  # local inputrack = find_pattern_by_name("INPUT")
  # INSPECT_CONFIG_MAP.append(create_inspect_config(item_id=3, dx=inputrack.pattern_width[0]/(inputrack.pattern_size[0]-1), dy=inputrack.pattern_width[1]/(inputrack.pattern_size[1]-1), rack_size=inputrack.pattern_size , description="Input Capture"))
  # # Fills the Landmark List with Projectrelated Data
  # # create_landmark(lm_id=0, marker_id=-1, marker_size=0.1, marker_type="aruco_7x7", capture_pos=p[0,0,0,0,0,0], init_frame=p[0,0,0,0,0,0], search_offset=[0,0,0], actual_frame=p[0,0,0,0,0,0], description="")
  # LANDMARK_MAP.append(create_landmark(lm_id=1, marker_id=3, marker_size=0.1, marker_type="aruco_7x7", capture_pos = F10_Cap_CF, init_frame=p[-0.617789, -0.065471, 0.07918, 0.020983, -0.012695, 1.512066], search_offset=[0.15, 0.15, 0.1], actual_frame=p[-0.617789, -0.065471, 0.07918, 0.020983, -0.012695, 1.512066], description="LM CF Lid"))
  # LANDMARK_MAP.append(create_landmark(lm_id=2, marker_id=-1, marker_size=0.0085, marker_type="aruco_4x4", capture_pos = F8_Cap_Cobas_LM, init_frame=p[0,0,0,0,0,0], search_offset=[0.15, 0.15, 0.1], actual_frame=POS_Z, description="LM Cobas Rack Detection"))
  # LANDMARK_MAP.append(create_landmark(lm_id=3, marker_id=0, marker_size=0.1, marker_type="aruco_7x7", capture_pos = F17_Cobas_Cap, init_frame=p[-0.667,-0.194,0.100,0,0,0], search_offset=[0.15, 0.15, 0.1], actual_frame=POS_Z, description="LM Cobas Cap"))
  # LANDMARK_MAP.append(create_landmark(lm_id=4, marker_id=4, marker_size=0.1, marker_type="aruco_7x7", capture_pos = F19_XN550_Cap, init_frame=p[0.124,-0.976,0.355,-0.008,0.025,3.131], search_offset=[0.15, 0.15, 0.1], actual_frame=p[0,0,0,0,0,0], description="LM XN550 Cap"))
  # LANDMARK_MAP.append(create_landmark(lm_id=5, marker_id=0, marker_size=0.1, marker_type="aruco_7x7", capture_pos = TestLMCap, init_frame=p[-0.49,-0.144,0.092,0,-0.008,0.001], search_offset=[0.15, 0.15, 0.1], actual_frame=POS_Z, description="LM Test"))
  # # Configuration of all movement related parameters
  # # create_movement(id=0, hh_approach=POS_Z, h_approach=POS_Z, approach=POS_Z, h_target=POS_Z, target=POS_Z, retract=POS_Z, h_retract=POS_Z, hh_retract=POS_Z, h_frame=POS_Z, frame=POS_Z, speed=1, acceleration=1, description="default")
  # MOVEMENT_MAP.append(create_movement(description="TestLMCap", frame=TestLMCap, actionlist=[ActionManipulator.MOVE_TO]))
  # MOVEMENT_MAP.append(create_movement(description="TestLM", frame=TestLM, actionlist=[ActionManipulator.PICK,ActionManipulator.PLACE],
  #         approach=p[0,0,0.1,0,0,0],
  #         retract=p[0,0,0.1,0,0,0]))
  # MOVEMENT_MAP.append(create_movement(description="Home - MOVE_TO", frame=F1_uLM_Home, actionlist=[ActionManipulator.MOVE_TO]))
  # MOVEMENT_MAP.append(create_movement(description="Input - PICK&PLACE", frame=F2_uLM_Input, actionlist=[ActionManipulator.PICK,ActionManipulator.PLACE],
  #         approach=p[0,0,0.1,0,0,0],
  #         retract=p[0,0,0.1,0,0,0]))
  # MOVEMENT_MAP.append(create_movement(description="Capture Input - MOVE_TO", frame=F3_Cap_Input, actionlist=[ActionManipulator.MOVE_TO]))
  # MOVEMENT_MAP.append(create_movement(description="BIN - PLACE", frame=F4_uLM_Bin, actionlist=[ActionManipulator.PLACE],
  #         approach=p[0,0,0.1,0,0,0],
  #         retract=p[0,0,0.1,0,0,0]))
  # MOVEMENT_MAP.append(create_movement(description="Gripper - Move To", frame=F5_uLM_Gripper, actionlist=[ActionManipulator.MOVE_TO],
  #         approach=p[0,0,0.1,0,0,0]))
  # MOVEMENT_MAP.append(create_movement(description="Gripper - Pick", frame=F5_uLM_Gripper, actionlist=[ActionManipulator.PICK],
  #         retract=p[0,0,0.1,0,0,0]))
  # MOVEMENT_MAP.append(create_movement(description="Gripper - Place", frame=F5_uLM_Gripper, actionlist=[ActionManipulator.PLACE],
  #         approach=p[0,0,0.1,0,0,0]))
  # MOVEMENT_MAP.append(create_movement(description="CobasRack Pick & Place", frame=F6_uLM_Cobas_R, actionlist=[ActionManipulator.PICK,ActionManipulator.PLACE],
  #         approach=p[0,0,0.1,0,0,0],
  #         target=p[0,0,0,0,0,d2r(90)],
  #         retract=p[0,0,0.1,0,0,0]))
  # MOVEMENT_MAP.append(create_movement(description="CobasMagazine Pick & Place", frame=F7_uLM_Coba_Mag, actionlist=[ActionManipulator.PICK,ActionManipulator.PLACE],
  #         approach=p[0,0,0.1,0,0,0],
  #         target=p[0,0,0,0,0,-d2r(90)],
  #         retract=p[0,0,0.1,0,0,0]))
  # MOVEMENT_MAP.append(create_movement(description="Capture Position Cobas Landmarks", frame=F8_Cap_Cobas_LM, actionlist=[ActionManipulator.MOVE_TO]))
  # MOVEMENT_MAP.append(create_movement(description="TaraMagazine - PICK & PLACE", frame=F9_uLM_Tara, actionlist=[ActionManipulator.PICK,ActionManipulator.PLACE],
  #         approach=p[0,0,0.13,0,0,0],
  #         target=p[0,0,0,0,0,-d2r(90)],
  #         retract=p[0,0,0.13,0,0,0]))
  # MOVEMENT_MAP.append(create_movement(description="Capture Position - Centrifuge LM", frame=F10_Cap_CF,actionlist=[ActionManipulator.MOVE_TO]))
  # MOVEMENT_MAP.append(create_movement(description="Pick and Place Racks - Centrifuge Lid", frame=F11_CF_PiPl, actionlist=[ActionManipulator.PICK,ActionManipulator.PLACE],
  #         approach=p[0,0,0.3,0,0,0],
  #         retract=p[0,0,0.3,0,0,0]))
  # MOVEMENT_MAP.append(create_movement(description="Pick and Place Samples - Centrifuge on uLM", frame=F12_uLM_CF_Mag, actionlist=[ActionManipulator.PICK,ActionManipulator.PLACE],
  #         approach=p[0,0,0.13,0,0,0],
  #         retract=p[0,0,0.13,0,0,0]
  #         ))
  # MOVEMENT_MAP.append(create_movement(description="Pick and Place Racks - Centrifuge on uLM", frame=F13_uLM_CF_R, actionlist=[ActionManipulator.PICK,ActionManipulator.PLACE],
  #         approach=p[0,0,0.15,0,0,0],
  #         retract=p[0,0,0.15,0,0,0]
  #         ))

  # MOVEMENT_MAP.append(create_movement(description="Pick and Place Samples XN550 Racks in Device", frame=F18_XN550_Input, actionlist=[ActionManipulator.PICK,ActionManipulator.PLACE],
  #         approach=p[0,0,0.1,0,0,0],
  #         target = p[0,0,0,0,0,d2r(90)],
  #         retract=p[0,0,0.1,0,0,0]
  #         ))
  # MOVEMENT_MAP.append(create_movement(description="Capture LM XN550", frame=F19_XN550_Cap, actionlist=[ActionManipulator.MOVE_TO]))
  # MOVEMENT_MAP.append(create_movement(description="Open XN550 Drawer ", frame=F20_XN550_Draw, actionlist=[ActionManipulator.DRAWER_OPEN],
  #         h_approach=p[0.07,0,0.1,0,0,0],
  #         approach=p[0,0,0.1,0,0,0],
  #         target = p[0,0,0,0,0,d2r(90)],
  #         retract=p[0.07,0,0,0,0,0],
  #         h_retract=p[0.07,0,0.1,0,0,0]
  #         ))
  # MOVEMENT_MAP.append(create_movement(description="Close XN550 Drawer ", frame=F20_XN550_Draw, actionlist=[ActionManipulator.DRAWER_CLOSE],
  #         h_approach=p[0.07,0,0.1,0,0,0],
  #         approach=p[0.07,0,0,0,0,0],
  #         target = p[0,0,0,0,0,d2r(90)],
  #         retract=p[0,0,0.1,0,0,0],
  #         h_retract=p[0.07,0,0.1,0,0,0]
  #         ))
  # MOVEMENT_MAP.append(create_movement(description="Push XN550 Button ", frame=F21_XN550_Btn, actionlist=[ActionManipulator.PUSH],
  #         approach=p[0,0,0.15,0,0,0],
  #         retract=p[0,0,0.15,0,0,0]
  #         ))
  # MOVEMENT_MAP.append(create_movement(description="Capture Position 2 Input", frame=F_Cap_Input2,actionlist=[ActionManipulator.MOVE_TO]))



  $ 19 "Script: SCRIPT Objects V0.1.script"
  #*****************************************************
  # customer          :   INTERNAL
  # project name      :
  #****************************************************
  # controller        :   UR
  # software          :   5.17.3
  #****************************************************
  # author            :   P. Koehnke
  # Copyright (c)     :   United Robotics Group
  #                       An der Riede 2
  #                       28816 Stuhr
  #                       Germany
  #****************************************************
  # description       :   object database
  # version:      	:   0.1
  # created           :   09.10.2024
  # updated           :
  #****************************************************
  # modifications     :
  #
  # date              :
  # name              :
  # reason            :
  #****************************************************

  def create_object_2(id=0, name="", type=0, dimension=struct(length=0, width=0, height=0, diameter=0), gripper_offset=p[0,0,0,0,0,0]):
      return struct(id=id, name=name, type=type, dimension=dimension, gripper_offset=gripper_offset)
  end

  OBJ = create_object_2()
  OBJs = make_list(0, create_object_2(), 50)

  OBJs.append(create_object_2(id=1, name="rack centrifuge", type=1, dimension=struct(length=0, width=0, height=0.106, diameter=0.020), gripper_offset=p[0,0,0.095,0,0,2.356]))
  OBJs.append(create_object_2(id=2, name="sample tube 1", type=2, dimension=struct(length=0, width=0, height=0.106, diameter=0.015), gripper_offset=p[0,0,0,0,0,0]))
  OBJs.append(create_object_2(id=3, name="rack sarstedt", type=3, dimension=struct(length=0, width=0, height=0.100, diameter=0.020), gripper_offset=p[0,0,0,0,0,0]))
  OBJs.append(create_object_2(id=4, name="Lab bottle", type=4, dimension=struct(length=0, width=0, height=0.100, diameter=0.030), gripper_offset=p[0,0,0.2,0,0,0]))
  OBJs.append(create_object_2(id=5, name="Vial", type=5, dimension=struct(length=0, width=0, height=0.100, diameter=0.0275), gripper_offset=p[0,0,0,0,0,0]))
  OBJs.append(create_object_2(id=6, name="Container", type=6, dimension=struct(length=0.0, width=0.0, height=0, diameter=0.0), gripper_offset=p[0,0,0,0,0,0]))
  OBJs.append(create_object_2(id=7, name="Target_container", type=7, dimension=struct(length=0.06, width=0.06, height=0.134, diameter=0.05), gripper_offset=p[0,0,0,0,0,0]))
  OBJs.append(create_object_2(id=8, name="Spatula", type=8, dimension=struct(length=0.03, width=0.03, height=0.23, diameter=0.05), gripper_offset=p[0,0,0,0,0,0]))
  OBJs.append(create_object_2(id=9, name="rack pipet", type=9, dimension=struct(length=0.03, width=0.03, height=0.23, diameter=0.05), gripper_offset=p[0,0,0,0,0,0]))

  def create_jig_2(id=0, name="", type=0, capacity=0, jig_offset=p[0,0,0,0,0,0]):
      # iformation about used jigs
      return struct(id=id, name=name, type=type, capacity=capacity, jig_offset=jig_offset)
  end

  JIG2 = create_jig_2()
  JIGs = make_list(0, create_jig_2(), 20)

  JIGs.append(create_jig_2(id=1, name="3FG", type=1, capacity=1, jig_offset=p[0,0,0,0,0,0]))
  JIGs.append(create_jig_2(id=2, name="jig input", type=2, capacity=1, jig_offset=p[0,0,0,0,0,-3.927]))
  JIGs.append(create_jig_2(id=3, name="jig output", type=3, capacity=1, jig_offset=p[0,0,0,0,0,0.78]))
  JIGs.append(create_jig_2(id=6, name="jig bin", type=6, capacity=1, jig_offset=p[0,0,0,0,0,0]))
  JIGs.append(create_jig_2(id=7, name="jig sarstedt racks", type=7, capacity=1, jig_offset=p[0,0,-0.02,0,0,0]))
  JIGs.append(create_jig_2(id=8, name="NoK Bin", type=8, capacity=1, jig_offset=p[0,0,0,0,0,0]))
  JIGs.append(create_jig_2(id=9, name="Pick bott jig", type=9, capacity=1, jig_offset=p[0,0,0,0,0,0]))
  JIGs.append(create_jig_2(id=10, name="Place bott jig", type=10, capacity=1, jig_offset=p[0,0,0,0,0,0]))
  JIGs.append(create_jig_2(id=11, name="bottle shake jig", type=11, capacity=1, jig_offset=p[0,0,0,0,0,0]))
  JIGs.append(create_jig_2(id=12, name="Pick Vial jig", type=12, capacity=1, jig_offset=p[0,0,0,0,0,0]))
  JIGs.append(create_jig_2(id=13, name="Place Vial jig", type=13, capacity=1, jig_offset=p[0,0,0,0,0,0]))
  JIGs.append(create_jig_2(id=14, name="Liquid transfer jig", type=14, capacity=1, jig_offset=p[0,0,0,0,0,0]))
  JIGs.append(create_jig_2(id=15, name="Pick station jig", type=15, capacity=1, jig_offset=p[0,0,0,0,0,0]))
  JIGs.append(create_jig_2(id=16, name="Place station jig", type=16, capacity=1, jig_offset=p[0,0,0,0,0,0]))
  JIGs.append(create_jig_2(id=17, name="Weigh station jig", type=17, capacity=1, jig_offset=p[0,0,0,0,0,0]))
  JIGs.append(create_jig_2(id=18, name="Pick station 1", type=18, capacity=1, jig_offset=p[0,0,0,0,0,0]))
  JIGs.append(create_jig_2(id=19, name="Pick station 2", type=19, capacity=1, jig_offset=p[0,0,0,0,0,0]))
  JIGs.append(create_jig_2(id=20, name="Pick station 3", type=20, capacity=1, jig_offset=p[0,0,0,0,0,0]))
  JIGs.append(create_jig_2(id=21, name="Tilt station jig", type=21, capacity=1, jig_offset=p[0,0,0,0,0,0]))
  $ 26 "Script: Powder_all.script"
  global SERVER_IP   = "192.168.12.139"
  global SERVER_PORT = 3002

  global container_id = 0
  global powder_id  = 0
  global bulk_density = 0
  global H          = 0
  global H_c          = 0
  global mouth_d     = 0
  global mouth_sh    = 0
  global length_c     = 0
  global diameter   = 0
  global empty_weight_g  = 0
  global volume_ml    = 0
  global shape_code   = 0
  global flow_code   = 0
  global shape = ""
  global Flowability = ""
  global full_weight_g = 0
  global cent_edge = 0
  global pick_2_base = 0.2 # distance from tcp to base of picking table
  global wall_thickness = 0.001

  def read_db_data():

    socket_open(SERVER_IP, SERVER_PORT)
    sleep(0.5)
    socket_send_string("GET_DATACODE_FLOATS")
    sleep(5)

    local fl = socket_read_ascii_float(14)
    socket_close()

    global container_id = fl[1]
    global powder_id = fl[2]
    global bulk_density = fl[3]
    global H          = fl[4]/1000
    global H_c          = fl[5]/1000
    global mouth_d     = fl[6]/1000
    global mouth_sh    = fl[7]/1000
    global length_c     = fl[8]/1000
    global diameter   = fl[9]/1000
    global empty_weight_g = fl[10]
    global volume_ml    = fl[11]
    global full_weight_g = fl[12]
    global flow_code   = fl[13]
    global shape_code   = fl[14]

  	if (flow_code == 1.0):
  	  global Flowability = "MEDIUM"
  	elif (flow_code == 2.0):
  	  global Flowability = "LOW"
  	else:
  	  global Flowability = "HIGH"
  	end

    if ( shape_code == 1.0):
  	shape = "cylindrical"
  	cent_edge =  diameter
    else:
  	shape = "cubical"
  	cent_edge =  length_c
    end

  end


  def send_picking_info(Pow_name, target_weight):
    socket_open(SERVER_IP, SERVER_PORT)
    cmd = "PICK:"+Pow_name+";"+to_str(target_weight)
    socket_send_string(cmd)
    sleep(0.1)
    socket_close()
  end

  #### POTS ####
  def tilt_send(angle):
  	socket_open("192.168.12.101", 80)
  	angle = 90.0 - angle
  	socket_send_string("Tilt,"+to_str(angle)+",0")
  	sync()
  	sleep(0.5)
  	socket_close()
  end

  def Motors_off():
  	socket_open("192.168.12.101", 80)
  	socket_send_string("Off,0,0")
  	sync()
  	sleep(0.5)
  	socket_close()
  end

  def Rotate():
  	socket_open("192.168.12.101", 80)
  	socket_send_string("FullRotation, 1, 2000")
  	sync()
  	sleep(0.5)
  	socket_close()
  end

  def CCW_Rotate():
  	socket_open("192.168.12.101", 80)
  	socket_send_string("FullRotation, -1, 2000")
  	sync()
  	sleep(0.5)
  	socket_close()
  end

  def tilt_to_home():
  	socket_open("192.168.12.101", 80)
  	socket_send_string("Home,0,0")
  	sync()
  	sleep(0.5)
  	socket_close()
  end
  #######
  def vibration_1():
  	set_analog_out(0,0.4)
  	sleep(1)
  	set_analog_out(0,0.0)
  	sleep(0)
  end

  def vibration_2():
  	set_analog_out(0,0.4)
  	sleep(0.8)
  	set_analog_out(0,0.0)
  	sleep(0.2)
  end

  def vibration_3():
  	set_analog_out(0,0.4)
  	sleep(0.5)
  	set_analog_out(0,0.0)
  	sleep(0.3)
  end

  def vibration_4():
  	set_analog_out(0,0.8)
  	sleep(0.6)
  	set_analog_out(0, 0.0)
  	sleep(0.5)
  end

  ##################

  global gear_2_holder = 0.018
  global gain_per_percent = 0.5
  global w_dosed_total = 0.0
  global last_scale = 0.0
  global tilt_angle_sent = 0.0
  global level = 0.0
  global target_g = 0.0
  global angle_max = 60
  global angle_min = 10
  global hinge_2_base = 0.0421
  global TCP_2_tip_x = 0.0047
  global spatula_len = 0.182
  global spatula_offset = p[TCP_2_tip_x,0,spatula_len,0,0,0]
  global SPATULA_L_VOL_ML = 5.0        # 1 teaspoon = 5 mL
  global SPATULA_M_VOL_ML = 1.25       # 1/4 teaspoon = 1.25 mL
  global SPATULA_S_VOL_ML = 0.15625    # 1/32 teaspoon = 0.15625 mL
  global SPATULA_FLAT_M_VOL_ML  = 2.2
  global SPATULA_FLAT_S_VOL_ML  = 1.2   #based on caluclations using rho = m/V
  global ry_deg_safe = 0
  global ry_deg = 0



  def clamp(x, lo, hi):
  	if(x<lo):
  		return lo
  	elif (x>hi):
  		return hi
  	else:
  		return x
  	end
  end

  def compute_level_percent(W_now, weight_value):   # W_now = container+powder, weight_value = live scale reading
      local delta = weight_value - last_scale

      if (delta < 0.0):
          delta = 0.0
      end

      global w_dosed_total = w_dosed_total + delta
      global last_scale = weight_value     # update the last scale reading

      local W_eff = W_now - w_dosed_total
      if (W_eff <  empty_weight_g):
          W_eff =  empty_weight_g
      end

      # Compute powder level %
      level = 100.0 * (W_eff -  empty_weight_g) / (full_weight_g -  empty_weight_g)

      # Clamp to 0–100
      level = clamp(level, 0, 100)
    textmsg("deb 1 = ", level)
      return level
  end

  def deg2rad(d):
  	return d*3.141592/180
  end

  def my_abs(val):
  	if (val<0):
  		return -val
  	else:
  		return val
  	end
  end

  def compute_tilt_deg(level_percent):
  	angle = angle_min + gain_per_percent*(100.0-level_percent)

    	textmsg("deb 2 = ", angle)
  	return clamp(angle, angle_min, angle_max)
  end

  def tilt(level_percentage):
  	new_angle = compute_tilt_deg(level_percentage)
  	global angle_rel = new_angle - tilt_angle_sent

  	if my_abs(angle_rel)>2.0:
  		tilt_send(new_angle)
  		global angle_deg = new_angle
  		global tilt_angle_sent = new_angle
  		global p_center_vertical = center_pose()
  		global p_center = updated_center_pose(p_center_vertical, angle_deg)
  	end

  	if (level_percentage<85.0):
  		tilt_send(angle_deg)
  	end
  end

  def compute_scoop_depth(level):
    return ((100.0-level)/100.0)*(H -mouth_sh )
  end

  def map_tilt_to_ry_deg(container_deg, level):

  	if (Flowability == "HIGH" or Flowability == "MEDIUM"):
  		global scoop_depth = compute_scoop_depth(level)
  		safe_scoop_pivot = (mouth_d  - spatula_depth)/(scoop_depth+mouth_sh )
  		global ry_deg_safe = asin(safe_scoop_pivot)
  		global ry_deg = 90-container_deg
  	else:
  		global scoop_depth = compute_scoop_depth(level)
  		safe_scoop_pivot = (mouth_d  - spatula_depth)/(scoop_depth+mouth_sh )
  		global ry_deg_safe = asin(safe_scoop_pivot)
  		global ry_deg = 90-container_deg
  	end
  	return [ry_deg_safe,ry_deg]
  end

  def get_scoop_weight(spatula, bulk_density):

  	local vol = 0

  	if (spatula == "spatula_L"):
  		vol = SPATULA_L_VOL_ML
  		global spatula_depth = 0.015
  		global spatula_mid   = 0.016
  		global spatula_ry    = 0.0

  	elif (spatula == "spatula_M"):
  		vol = SPATULA_M_VOL_ML
  		global spatula_depth = 0.010
  		global spatula_mid   = 0.0105
  		global spatula_ry    = 0.0

  	elif (spatula == "spatula_S"):
  		vol = SPATULA_S_VOL_ML
  		global spatula_depth = 0.008
  		global spatula_mid   = 0.0063
  		global spatula_ry    = 0.0

  	elif (spatula == "spatula_flat_M"):
  		vol = SPATULA_FLAT_M_VOL_ML
  		global spatula_depth = 0.001
  		global spatula_mid   = 0.002
  		global spatula_ry    = 10.0

  	elif (spatula == "spatula_flat_S"):
  		vol = SPATULA_FLAT_S_VOL_ML
  		global spatula_depth = 0.005
  		global spatula_mid   = 0.016
  		global spatula_ry    = 2.0

  	else:
  		textmsg("Unknown spatula type")
  		return 0.0
  	end
  	global target_g = vol * bulk_density
  	return target_g

  end

  def select_spatula(Flowability, level, diff, bulk_density, mouth_d ):

      local k = 1.1

      global powder_height = (H  - mouth_sh ) * level/100

      # =====================================================
      # LOW FLOWABILITY
      # =====================================================
      if (Flowability == "LOW"):

          local gFM = get_scoop_weight("spatula_flat_M", bulk_density)

          local level_ok_FM = (spatula_mid * 2 < powder_height)
          local diff_ok_FM  = (diff > k * gFM)

          local flatM_ok = level_ok_FM and diff_ok_FM

          if (flatM_ok):
              return "spatula_flat_M"
          else:
              return "spatula_flat_S"
          end

      end


      # =====================================================
      # LARGE
      # =====================================================
      local gL = get_scoop_weight("spatula_L", bulk_density)

      local mouth_ok_L = (mouth_d  >= 0.05)
      local level_ok_L = (spatula_mid * 2 < powder_height)
      local diff_ok_L  = (diff > k * gL)

      local large_ok = mouth_ok_L and level_ok_L and diff_ok_L


      # =====================================================
      # MEDIUM
      # =====================================================
      local gM = get_scoop_weight("spatula_M", bulk_density)

      local level_ok_M = (spatula_mid * 2 < powder_height)
      local diff_ok_M  = (diff > k * gM)

      local medium_ok = level_ok_M and diff_ok_M


      # =====================================================
      # FINAL SELECTION
      # =====================================================
      if (large_ok):
          return "spatula_L"

      elif (medium_ok):
          return "spatula_M"

      else:
          return "spatula_S"
      end

  end

  def after_scoop():
  	tilt_send(angle_deg)
  	sleep(0.5)
  	movel(lifted_pose, a=0.05, v=0.2)
  	movel(tilted_pose_in_base2, a=0.05, v=0.2)
  	set_analog_out(0,0.4)
  	movel(pose_trans(tilted_pose_in_base2, p[0,0,0,0,0,2.0]), a=0.05, v=0.2)
  	set_analog_out(0,0.0)
  	movel(lifted_pose, a=0.05, v=0.2)
  	tilt_to_home()
  end

  def center_pose():
  	global p_translated = container_place
  	#global p_translated = pots_axis_temp

  	#cx = p_translated[0]
  	#cy = p_translated[1]
  	#cz = p_translated[2]

  	global p_center_vertical_temp = pose_trans(p_translated, p[0,0,0, deg2rad(90), 0, 0])
  	cx = p_center_vertical_temp[0]
  	cy = p_center_vertical_temp[1]
  	cz = p_center_vertical_temp[2]
  	#rx = p_center_vertical_temp[3]
  	#ry = p_center_vertical_temp[4]
  	rz = p_center_vertical_temp[5]

  	global p_center_vertical_temp = p[cx,cy,cz, 0, 0, rz]
  	trans_rel = p[0,0,-pick_2_base+H,0,0,0]
  	global p_center_vertical =  pose_trans(p_center_vertical_temp, trans_rel)
  	return p_center_vertical
  end

  def updated_center_pose(p_center_vertical, angle_deg):
  	hinge_pose = pose_trans(p_center_vertical, p[0,0,-hinge_2_base-gear_2_holder-H ,0,0,0])
  	local_rel = pose_trans(pose_inv(hinge_pose), p_center_vertical)

  	rot_tilt = p[0,0,0, -deg2rad(angle_deg),0,0]
  	local_rel_tilted = pose_trans(rot_tilt, local_rel)

  	global p_center = pose_trans(hinge_pose, local_rel_tilted)
  	return p_center
  end

  def scoop_powder(p_center):
  	vibration_voltage = 0.4
  	vibration_time = 3.0
  	global scoop_radius_default = 0.0


  	scoop_radius_default = mouth_d /2 - spatula_depth
  	scoop_safe_entry_pose = pose_trans(p_center, p[-TCP_2_tip_x,0,spatula_len+0.05,0,0,0])
  	scoop_entry_pose = pose_trans(p_center, p[-TCP_2_tip_x,0,spatula_len,0,0,0])

  	movel(scoop_safe_entry_pose, a=0.1, v=0.25)
  	movel(scoop_entry_pose, a=0.1, v=0.25)

  	scoop_start_rel_int = p[0, 0, -mouth_sh , 0, 0, 0]
  	scoop_start_pose_int = pose_trans(scoop_entry_pose, scoop_start_rel_int)

  	movel(scoop_start_pose_int, a=0.1, v=0.25)

  	if (spatula_mid * 2 < powder_height and spatula == "spatula_M" or spatula == "spatula_L"):

  		global total_depth = mouth_sh + scoop_depth + spatula_mid
  		global total_depth = clamp(total_depth, 0, H - spatula_mid)
  		scoop_start_rel = p[scoop_radius_default, 0, -total_depth, 0, 0, 0]

  		rot_mid = p[0, 0, 0, 0, 0, 0.785]
  		rot_end = p[0, 0, 0, 0, 0, 1.5708]

  		scoop_via_rel = pose_trans(rot_mid, scoop_start_rel)
  		scoop_end_rel = pose_trans(rot_end, scoop_start_rel)

  		scoop_start_pose = pose_trans(scoop_entry_pose, scoop_start_rel)
  		scoop_via_pose = pose_trans(scoop_entry_pose, scoop_via_rel)
  		scoop_end_pose = pose_trans(scoop_entry_pose, scoop_end_rel)

  		movel(scoop_start_pose, a=0.5, v=0.3)

  		if (level<90.0):
  			Rotate()
  		end

  		movec(scoop_via_pose, scoop_end_pose, a=0.03, v=0.02)
  		sleep(1.0)
  		#local ry_deg = map_tilt_to_ry_deg(angle_deg,level)
  		local ry_result = map_tilt_to_ry_deg(angle_deg,level)
  		global ry_safe = ry_result[0]
  		global ry = deg2rad(ry_result[1])

  		# safe_retention
  		local pivot_pose = pose_trans(scoop_end_pose, p[0,0,total_depth-spatula_len,0,0,0])
  		local end_rel = pose_trans(pose_inv(pivot_pose), scoop_end_pose)
  		local end_rel_tilted = pose_trans(end_rel, p[0, 0, 0, 0, ry_safe, 0])
  		global tilted_pose_in_base = pose_trans(pivot_pose, p[0,0,0,end_rel_tilted[3],end_rel_tilted[4], end_rel_tilted[5]])
  		global tilted_pose_in_base = pose_trans(tilted_pose_in_base, p[0, 0, spatula_len-total_depth, 0, 0, 0])
  		# sptula pivoted around the container rim of the mouth at ry_safe
  		movel(tilted_pose_in_base, a=0.03, v=0.1)

  		#popup("is the spatula crashing at front? ", blocking = True)
  		# safe_retention_above
  		# calculate x , z movements

  		global safe_x = sin(ry_safe)*(scoop_depth - (mouth_d -spatula_depth)/tan(90-ry_safe/2))
  		global safe_z = cos(ry_safe)*(scoop_depth - (mouth_d -spatula_depth)/tan(90-ry_safe/2))

  		local safe_up = pose_trans(tilted_pose_in_base, p[-safe_x,0,safe_z,0,0,0])
  		movel(safe_up, a=0.03, v=0.1)

  		#popup("is the spatula crashing at neck? ", blocking = True)

  		# full exit step by step
  		#local alpha = atan(2*mouth_sh /mouth_d )

  		#global cent_pose_cont_x = sin(ry_safe)*(scoop_depth - (mouth_d -spatula_depth)/tan(90-ry_safe/2))
  		#global cent_pose_cont_z = cos(ry_safe)*(scoop_depth+mouth_sh  - (mouth_d -spatula_depth)/tan(90-ry_safe/2))
  		#local cent_pose_cont = pose_trans(safe_up, p[])

  		# full exit
  		local pivot_pose2 = pose_trans(tilted_pose_in_base, p[0,0,total_depth-spatula_len,0,0,0])
  		local end_rel2 = pose_trans(pose_inv(pivot_pose2), tilted_pose_in_base)
  		#popup("is the spatula crashing front? ", blocking = True)
  		local end_rel_tilted2 = pose_trans(end_rel2, p[0, 0, 0, 0, ry-ry_safe, 0])
  		global tilted_pose_in_base2 = pose_trans(pivot_pose2, p[0,0,0,end_rel_tilted2[3],end_rel_tilted2[4], end_rel_tilted2[5]])
  		global tilted_pose_in_base2 = pose_trans(tilted_pose_in_base2, p[-TCP_2_tip_x, 0, spatula_len-scoop_radius_default-spatula_mid, 0, 0, 0])
  		# spaula exited at center of the mouth at ry
  		movel(tilted_pose_in_base2, a=0.03, v=0.1)
  		#popup("is the spatula crashing at mouth? ", blocking = True)

  	else : # emptying logic
  		spatula_base = pose_trans(scoop_entry_pose, p[0, 0, -H, 0, 0, 0])
  		local pivot_pose = pose_trans(scoop_entry_pose, p[0,0,-spatula_len,0,0,0])
  		# tilt inwards
  		global in_angle = atan((cent_edge-spatula_depth)/(2*H))
  		spatula_tilt_rel = pose_trans(pose_inv(pivot_pose), spatula_base)

  		spatula_tilt = pose_trans(spatula_tilt_rel, p[0, 0, 0, in_angle, 0, 0])
  		global tilted_pose = pose_trans(pivot_pose, p[0,0,0,spatula_tilt[3],spatula_tilt[4], spatula_tilt[5]])

  		global tilted_pose = pose_trans(tilted_pose, p[0,0,spatula_len-H,0,0,0])

  		movel(tilted_pose,a=0.1, v=0.25)
  		Rotate()

  		rot_mid = p[0, 0, 0, 0, 0, 0.785]
  		rot_end = p[0, 0, 0, 0, 0, 1.5708]

  		scoop_via_rel = pose_trans(tilted_pose, rot_mid)
  		scoop_end_rel = pose_trans(tilted_pose, rot_end)

  		movec(scoop_via_rel, scoop_end_rel, a=0.03, v=0.02)
  		popup("is the spatula crashing front? ", blocking = True)

  		scoop_via_pose = pose_trans(pivot_pose, scoop_via_rel)
  		scoop_end_pose = pose_trans(pivot_pose, scoop_end_rel)

  		#movec(scoop_via_pose, scoop_end_pose, a=0.03, v=0.02)
  		popup("is the spatula crashing front? ", blocking = True)
  		local ry_result = map_tilt_to_ry_deg(angle_deg,level)
  		global ry_safe = ry_result[0]
  		global ry = deg2rad(ry_result[1])

  		# full exit
  		#local pivot_pose2 = pose_trans(scoop_entry_pose, p[0,0,-spatula_len,0,0,0])
  		local end_rel2 = pose_trans(pose_inv(pivot_pose), scoop_end_pose)
  		popup("is the spatula crashing front? ", blocking = True)
  		local end_rel_tilted2 = pose_trans(end_rel2, p[0, 0, 0, 0, ry, 0])
  		global tilted_pose_in_base2 = pose_trans(pivot_pose, p[0,0,0,end_rel_tilted2[3],end_rel_tilted2[4], end_rel_tilted2[5]])
  		global tilted_pose_in_base2 = pose_trans(tilted_pose_in_base2, p[0, 0, spatula_len, 0, 0, 0])
  		# sptula exited at center of the mouth at ry
  		movel(tilted_pose_in_base2, a=0.03, v=0.1)
  		popup("is the spatula crashing at mouth? ", blocking = True)
  	end

  	if (spatula=="spatula_flat_S" or spatula=="spatula_S"):
  		vibration_3()
  	elif (spatula == "spatula_M"):
  		vibration_4()
  	else:
  		set_analog_out(0, vibration_voltage)
  	end

  	# remove excess
  	local pivot_pose_level = pose_trans(tilted_pose_in_base2, p[0,0,-spatula_len,0,0,0])
  	local end_rel_level = pose_trans(pose_inv(pivot_pose_level), tilted_pose_in_base2)
  	#local ry_level = ry/1.5
  	local ry_level = deg2rad(15)
  	local end_rel_tilted_level = pose_trans(end_rel_level, p[0, 0, 0, 0, -ry_level, 0])
  	local end_rel_tilted_level2 = pose_trans(pivot_pose_level, p[0, 0, 0,end_rel_tilted_level[3],end_rel_tilted_level[4], end_rel_tilted_level[5]])
  	local end_rel_tilted_level2 = pose_trans(end_rel_tilted_level2, p[0,0,spatula_len,0,0,0])
  	movel(end_rel_tilted_level2, a=0.03, v=0.1)

  	movel(tilted_pose_in_base2, a=0.03, v=0.1)
  	set_analog_out(0, 0.0)
  	#popup("safe out + moving towards beaker", title = "Pause", blocking = True)
  	global lifted_pose = pose_trans(tilted_pose_in_base2, p[-0.04,0,0.04,0,0,0]) # safety distance away from the container

  	movel(lifted_pose, a=0.03, v=0.1)
  	CCW_Rotate()
  end

  def auto_tilt_and_scoop(W_now, target_weight, weight_value):
  	global level = compute_level_percent(W_now, weight_value)

  	global spatula = select_spatula(Flowability, level, diff, bulk_density, mouth_d )
  	textmsg("deb 4 8 = ", spatula)
  	#global target_g = get_scoop_weight(spatula, bulk_density)

    	#textmsg("deb 4 = ", target_g)
  	#send_scoop_target_info()

  	global scoop_depth = compute_scoop_depth(level)

    	textmsg("deb 5 = ", scoop_depth)
  	tilt_to_home()
  	sleep(0.5)
  	tilt(level)
  	sleep(1.5)
    	#popup("is the pots tilted? ", blocking = True)
    	#textmsg("deb 6 = ", p_center)
  	scoop_powder(p_center)

    	textmsg("deb 7 - sucess")
  end
  $ 27 "Script: Weight_scale_socket_s.script"
  global s_depth = 0
  global s_length =0
  global s_volume = 0
  global ry_theta  = 0

  def get_weight():
  	socket_open(SERVER_IP,SERVER_PORT)
  	sleep(0.2)
  	textmsg("socket opened successfully!")
  	socket_send_string("GET_WEIGHT")
  	sleep(0.2)
  	sync()
  	sleep(0.2)
  	receiveFromServ = socket_read_ascii_float(6)
  	sleep(1)
  	#while (receiveFromServ[0] <1):
  		#receiveFromServ = socket_read_ascii_float(1)
  		#sleep(1)
  		#textmsg("retrying read:", receiveFromServ)
  	#end
  	textmsg("Received weight:", receiveFromServ[1])
  	sleep(0.2)
  	socket_close()
  	sleep(0.2)
  	return receiveFromServ[1]
  end

  def tare_scale():
  	socket_open(SERVER_IP,SERVER_PORT)
  	socket_send_string("TARE")
  	sleep(2)
  	socket_close()
  end

  def zero_scale():
  	socket_open(SERVER_IP,SERVER_PORT)
  	socket_send_string("ZERO")
  	sleep(0.5)
  	socket_close()
  end

  def log_weight():
  	socket_open(SERVER_IP,SERVER_PORT)
  	socket_send_string("LOG_WEIGHT")
  	sleep(0.5)
  	socket_close()
  end

  def send_target_info():
  	socket_open(SERVER_IP,SERVER_PORT)
  	socket_send_string("SET_TARGET:" + to_str(target_weight))
  	sleep(0.2)
  	socket_close()
  end
  def send_powder_info():
  	socket_open(SERVER_IP,SERVER_PORT)
  	socket_send_string("SET_POWDER:" + Pow_name)
  	sleep(0.2)
  	socket_close()
  end
  def send_spatula_info():
  	socket_open(SERVER_IP,SERVER_PORT)
  	socket_send_string("SET_SPATULA:" + spatula)
  	#sleep(1)

  	#local fl = socket_read_ascii_float(4)
    	#socket_close()

    	#global s_depth = fl[1]
    	#global s_length = fl[2]
   	#global s_volume = fl[3]
   	#global ry_theta  = fl[4]
  	sleep(0.2)

  end

  def send_level_info():
  	socket_open(SERVER_IP,SERVER_PORT)
  	socket_send_string("SET_LEVEL:" + to_str(level))
  	sleep(0.2)
  	socket_close()
  end
  def send_weight_info():
    socket_open(SERVER_IP, SERVER_PORT)
    #rq_open_and_wait()
    cmd = "GET_CONT_WEIGHT"
    socket_send_string(cmd)
    sync()
    sleep(0.5)
    receiveFromSer = socket_read_ascii_float(1)
    socket_close()
    return receiveFromSer[1]
  end

  $ 28 "BeforeStarts"
  $ 29 "uLM"
  $ 30 "CMD_Stop≔ False "
  global CMD_Stop=  False
  $ 31 "CMD_Abort≔ False "
  global CMD_Abort=  False
  $ 32 "CMD_Clear≔ False "
  global CMD_Clear=  False
  $ 33 "STATE≔1"
  global STATE=1
  $ 34 "STATE_Info≔''"
  global STATE_Info=""
  $ 35 "ARM_Referenced≔ False "
  global ARM_Referenced=  False
  $ 36 "zero_ftsensor()"
  zero_ftsensor()
  $ 37 "poses init"
  $ 38 "PSE_A≔p[0,0,0,0,0,0]"
  global PSE_A=p[0,0,0,0,0,0]
  $ 39 "PSE_A_H≔p[0,0,0,0,0,0]"
  global PSE_A_H=p[0,0,0,0,0,0]
  $ 40 "PSE_R≔p[0,0,0,0,0,0]"
  global PSE_R=p[0,0,0,0,0,0]
  $ 41 "PSE_R_H≔p[0,0,0,0,0,0]"
  global PSE_R_H=p[0,0,0,0,0,0]
  $ 42 "PSE_T≔p[0,0,0,0,0,0]"
  global PSE_T=p[0,0,0,0,0,0]
  $ 43 "PSE_T_H≔p[0,0,0,0,0,0]"
  global PSE_T_H=p[0,0,0,0,0,0]
  $ 44 "PSE_C_E≔p[0,0,0,0,0,0]"
  global PSE_C_E=p[0,0,0,0,0,0]
  $ 45 "PSE_C_H≔p[0,0,0,0,0,0]"
  global PSE_C_H=p[0,0,0,0,0,0]
  $ 46 "PSE_C_S≔p[0,0,0,0,0,0]"
  global PSE_C_S=p[0,0,0,0,0,0]
  $ 47 "init_home_by_cartesian_pose(p[0,-0.400,0.300,0,0,0])"
  init_home_by_cartesian_pose(p[0,-0.400,0.300,0,0,0])
  $ 48 "Clearing"
  $ 49 "reset_error()"
  reset_error()
  $ 50 "reset_warning()"
  reset_warning()
  $ 51 "uGo"
  $ 53 "ugo_init( True ,'http://192.168.12.120:10001')"
  ugo_init(  True  ,"http://192.168.12.120:10001")
  $ 54 "ugo_update_outputs()"
  ugo_update_outputs()
  $ 55 "App"
  $ 56 "'ADD APPLICATION SPECIFIC COMMANDS'"
  # 'ADD APPLICATION SPECIFIC COMMANDS'
  $ 57 "Tools"
  $ 58 "OBJ_Picked≔gripper_has_object()"
  global OBJ_Picked=gripper_has_object()
  $ 59 "If OBJ_Picked"
  if (OBJ_Picked):
    # begin: URCap Program Node
    #   Source: Robotiq_Grippers, 3.17.0.105337, Robotiq Inc.
    #   Type: Gripper Activate
    $ 60 "Gripper Activate"

    kill rq_gripper_communication_thread
    rq_gripper_communication_thread_started = False
    rq_close_gripper_socket("1")
    rq_close_gripper_socket("2")
    rq_close_gripper_socket("3")
    rq_close_gripper_socket("4")

    rq_init_comm_if_connected(9, "1")
    rq_init_comm_if_connected(2, "2")
    rq_init_comm_if_connected(3, "3")
    rq_init_comm_if_connected(4, "4")
    rq_print_connected_grippers()
    rq_gripper_communication_thread = run rq_gripper_communication()

    while(not rq_gripper_communication_thread_started):
        sleep(0.008)
    end

    rq_set_max_current_for_all_grippers()

    reset_and_activate = False

    rq_activate_all_grippers(False)
    # end: URCap Program Node
  else:
    $ 61 "Else" "noBreak"
    # begin: URCap Program Node
    #   Source: Robotiq_Grippers, 3.17.0.105337, Robotiq Inc.
    #   Type: Gripper Activate
    $ 62 "Gripper Reset and Activate"

    kill rq_gripper_communication_thread
    rq_gripper_communication_thread_started = False
    rq_close_gripper_socket("1")
    rq_close_gripper_socket("2")
    rq_close_gripper_socket("3")
    rq_close_gripper_socket("4")

    rq_init_comm_if_connected(9, "1")
    rq_init_comm_if_connected(2, "2")
    rq_init_comm_if_connected(3, "3")
    rq_init_comm_if_connected(4, "4")
    rq_print_connected_grippers()
    rq_gripper_communication_thread = run rq_gripper_communication()

    while(not rq_gripper_communication_thread_started):
        sleep(0.008)
    end

    rq_set_max_current_for_all_grippers()

    reset_and_activate = True

    rq_activate_all_grippers(True)
    # end: URCap Program Node
  end
  $ 63 "zero_ftsensor()"
  zero_ftsensor()
  $ 64 "EXTT"
  $ 65 "Set GRP_3F_Enable=Off"
  set_standard_digital_out(4, False)
  $ 66 "Set BarcodeTrigger=Off"
  set_standard_digital_out(6, False)
  $ 67 "Set GRP_3F_Decap=Off"
  set_standard_digital_out(3, False)
  $ 68 "Set GRP_3F_Cap=Off"
  set_standard_digital_out(2, False)
  $ 69 "Set GRP_3F_Open=Off"
  set_standard_digital_out(5, False)
  $ 70 "PSE_T≔get_tool_free_pose(dir=[0,0,0.150], move_in_base_frame=True)"
  global PSE_T=get_tool_free_pose(dir=[0,0,0.150], move_in_base_frame=True)
  $ 71 "If is_reachable(Base_const, [PSE_T])"
  if (is_reachable(p[0.0,0.0,0.0,0.0,0.0,0.0], [PSE_T])):
    $ 72 "MoveL"
    $ 73 "PSE_T" "breakAfter"
    movel(PSE_T, a=1.2, v=0.15)
  end
  $ 75 "powder dispensing variable init"
  $ 76 "Start_thread≔ False "
  global Start_thread=  False
  $ 77 "vib_thread≔ False "
  global vib_thread=  False
  $ 78 "QR assignment init"
  $ 79 "d_cc≔0.06"
  global d_cc=0.06
  $ 81 "kp≔0.0015"
  global kp=0.0015
  $ 82 "ki≔0.0001"
  global ki=0.0001
  $ 83 "kd≔0.01"
  global kd=0.01
  $ 84 "dt≔0.03"
  global dt=0.03
  $ 85 "Integral_error≔0"
  global Integral_error=0
  $ 86 "current_error≔0"
  global current_error=0
  $ 87 "previous_error≔0"
  global previous_error=0
  $ 88 "tilt_increment≔0"
  global tilt_increment=0
  $ 89 "tilt_angle≔0"
  global tilt_angle=0
  $ 90 "diff≔0"
  global diff=0
  $ 91 "current_pose≔get_actual_tcp_pose()"
  global current_pose= get_actual_tcp_pose ()
  $ 92 "Relative_trans≔p[0, 0, -0.035, 0, 0, 0]"
  global Relative_trans=p[0, 0, -0.035, 0, 0, 0]
  $ 96 "tilt_to_home()"
  tilt_to_home()
  $ 97 "switch_spat_M≔ True "
  global switch_spat_M=  True
  $ 98 "switch_spat_S≔ True "
  global switch_spat_S=  True
  $ 99 "switch_spat_F_M≔ True "
  global switch_spat_F_M=  True
  $ 100 "switch_spat_F_S≔ True "
  global switch_spat_F_S=  True
  $ 101 "last_scale≔0"
  global last_scale=0
  $ 793 "Thread_1"
  thread Thread_1():
    while (True):
      $ 794 "If Start_thread≟ True "
      if (Start_thread ==   True  ):
        $ 795 "weight_value≔get_weight()"
        global weight_value=get_weight()
        $ 796 "Wait: 0.2"
        sleep(0.2)
        $ 797 "sync()"
        sync()
      end
      $ 798 "sync()"
      sync()
    end
  end
  threadId_Thread_1 = run Thread_1()
  $ 799 "Thread_2"
  thread Thread_2():
    while (True):
      $ 800 "Loop vib_thread≟ True "
      thread Thread_while_800():
        while (True):
          $ 801 "diff≔target_weight-weight_value"
          global diff=target_weight-weight_value
          $ 802 "If diff>0.02 and spatula≠'spatula_flat_S'"
          global thread_flag_802=0
          thread Thread_if_802():
            $ 804 "Set AO[0]=4.0"
            set_standard_analog_out(0, 0.4)
            thread_flag_802 = 1
          end
          if (diff>0.02  and  spatula != "spatula_flat_S"):
            global thread_handler_802=run Thread_if_802()
            while (thread_flag_802 == 0):
              if not(diff>0.02  and  spatula != "spatula_flat_S"):
                kill thread_handler_802
                thread_flag_802 = 2
              else:
                sync()
              end
            end
          else:
            thread_flag_802 = 2
          end
          if (thread_flag_802 == 2):
            $ 805 "ElseIf diff>0.02 and spatula≟'spatula_flat_S'"
            if (diff>0.02 and spatula == "spatula_flat_S"):
              $ 806 "vibration_3()"
              vibration_3()
            else:
              $ 807 "ElseIf diff≤0.03"
              global thread_flag_807=0
              thread Thread_if_807():
                $ 808 "vibration_2()"
                vibration_2()
                thread_flag_807 = 1
              end
              if (diff <= 0.03):
                global thread_handler_807=run Thread_if_807()
                while (thread_flag_807 == 0):
                  if not(diff <= 0.03):
                    kill thread_handler_807
                    thread_flag_807 = 2
                  else:
                    sync()
                  end
                end
              else:
                thread_flag_807 = 2
              end
              if (thread_flag_807 == 2):
                $ 813 "Else" "noBreak"
                $ 814 "Set AO[0]=0.0"
                set_standard_analog_out(0, 0.0)
              end
            end
          end
        end
      end
      if (vib_thread ==   True  ):
        global thread_handler_800=run Thread_while_800()
        while (vib_thread ==   True  ):
          sync()
        end
        kill thread_handler_800
      end
      $ 815 "sync()"
      sync()
    end
  end
  threadId_Thread_2 = run Thread_2()
  while (True):
    $ 102 "Robot Program"
    $ 103 "MAIN"
    $ 104 "command_manager(external_control='uGO', cond_suspend=(ITM_Manipulated and AMR_AtTarget and AMR_Charging and AMR_Battery<40), cond_unsuspend=(AMR_Battery≟60))"
    command_manager(external_control="uGO", cond_suspend=(ITM_Manipulated  and  AMR_AtTarget  and  AMR_Charging  and  AMR_Battery<40), cond_unsuspend=(AMR_Battery == 60))
    $ 105 "log_state(STATE_Info)"
    log_state(STATE_Info)
    $ 106 "Switch STATE"
    switch_1 = STATE
    $ 107 "Case 1"
    if (1 == switch_1):
      $ 108 "Stopping"
      $ 109 "STATE_Info≔'Stopping'"
      global STATE_Info="Stopping"
      $ 110 "end_freedrive_mode()"
      end_freedrive_mode()
      $ 111 "Set"
      set_tcp(p[0.0,0.0,0.161,3.1415,0.0,0.0])
      $ 112 "PSE_T≔get_tool_free_pose(dir=[0,0,0.150], move_in_base_frame=True)"
      global PSE_T=get_tool_free_pose(dir=[0,0,0.150], move_in_base_frame=True)
      $ 113 "If is_reachable(Base_const, [PSE_T])"
      if (is_reachable(p[0.0,0.0,0.0,0.0,0.0,0.0], [PSE_T])):
        $ 114 "MoveL"
        $ 115 "PSE_T" "breakAfter"
        movel(PSE_T, a=1.2, v=0.15)
      end
      $ 116 "do_transition(keep_rxry=OBJ_Picked, r=0)"
      do_transition(keep_rxry=OBJ_Picked, r=0)
      $ 125 "Call Sub_AMR_MiR_V3"
      Sub_AMR_MiR_V3()
      $ 126 "If stopping() and AMR_Done"
      if (stopping()  and  AMR_Done):
        $ 127 "STATE≔2"
        global STATE=2
        $ 128 "ugo_update_outputs()"
        ugo_update_outputs()
      end
    elif (2 == switch_1):
      $ 129 "Case 2"
      $ 130 "Stopped"
      $ 131 "STATE_Info≔'Stopped'"
      global STATE_Info="Stopped"
      $ 132 "Call Sub_AMR_MiR_V3"
      Sub_AMR_MiR_V3()
      $ 133 "If CMD_Reset  or PB_Start"
      if (CMD_Reset   or  get_standard_digital_in(0)):
        $ 134 "STATE≔3"
        global STATE=3
        $ 135 "ugo_update_outputs()"
        ugo_update_outputs()
      end
    elif (3 == switch_1):
      $ 136 "Case 3"
      $ 137 " Resetting"
      $ 138 "STATE_Info≔'Resetting'"
      global STATE_Info="Resetting"
      $ 139 "uML"
      $ 140 "reset_error()"
      reset_error()
      $ 141 "reset_warning()"
      reset_warning()
      $ 142 "PROCESS_Step≔0"
      global PROCESS_Step=0
      $ 143 "PROCESS_Info≔''"
      global PROCESS_Info=""
      $ 144 "ARM_Referenced≔ False "
      global ARM_Referenced=  False
      $ 145 "WRK_Done≔ False "
      global WRK_Done=  False
      $ 146 "ITM_Prepared≔ False "
      global ITM_Prepared=  False
      $ 147 "ITM_Manipulated≔ False "
      global ITM_Manipulated=  False
      $ 148 "STP≔0"
      global STP=0
      $ 149 "Action≔0"
      global Action=0
      $ 150 "Action_Info≔''"
      global Action_Info=""
      $ 151 "ITM_ID≔0"
      global ITM_ID=0
      $ 152 "JIG≔0"
      global JIG=0
      $ 153 "JIG_Slot≔0"
      global JIG_Slot=0
      $ 154 "Task_info≔''"
      global Task_info=""
      $ 155 "Set"
      set_tcp(p[0.0,0.0,0.161,3.1415,0.0,0.0])
      $ 156 "App"
      $ 157 "'ADD APPLICATION SPECIFIC COMMANDS'"
      # 'ADD APPLICATION SPECIFIC COMMANDS'
      $ 158 "OBJ_Type≔0"
      global OBJ_Type=0
      $ 159 "OBJ_Nbr≔0"
      global OBJ_Nbr=0
      $ 160 "If CNT_Rack_Output≥50"
      if (CNT_Rack_Output >= 50):
        $ 161 "CNT_Rack_Output≔0"
        global CNT_Rack_Output=0
      end
      $ 162 "TASK≔struct(ID=0, NAVI=struct(target=0, footprint=0, protectiveOff=0, dock=0), WORK=struct(ITM_ID_Src=0, JIG_ID_Src=0, OBJ_Nbr_Src=0, ACT_Src=0, ITM_ID_Tgt=0, JIG_ID_Tgt=0, OBJ_Nbr_Tgt=0, ACT_Tgt=0, OBJ_Type=0))"
      global TASK=struct(ID=0, NAVI=struct(target=0, footprint=0, protectiveOff=0, dock=0), WORK=struct(ITM_ID_Src=0, JIG_ID_Src=0, OBJ_Nbr_Src=0, ACT_Src=0, ITM_ID_Tgt=0, JIG_ID_Tgt=0, OBJ_Nbr_Tgt=0, ACT_Tgt=0, OBJ_Type=0))
      $ 163 "Call Sub_AMR_MiR_V3"
      Sub_AMR_MiR_V3()
      $ 164 "If resetting() and AMR_Done"
      if (resetting()  and  AMR_Done):
        $ 165 "STATE≔4"
        global STATE=4
        $ 166 "ugo_update_outputs()"
        ugo_update_outputs()
      end
    elif (4 == switch_1):
      $ 167 "Case 4"
      $ 168 "Idle"
      $ 169 "STATE_Info≔'Idle'"
      global STATE_Info="Idle"
      $ 170 "If CMD_Start"
      if (CMD_Start):
        $ 171 "STATE≔5"
        global STATE=5
        $ 172 "ugo_update_outputs()"
        ugo_update_outputs()
      end
    elif (5 == switch_1):
      $ 173 "Case 5"
      $ 174 "Starting"
      $ 175 "STATE_Info≔'Starting'"
      global STATE_Info="Starting"
      $ 176 "'ADD COMMANDS WHAT TO START WITH'"
      # 'ADD COMMANDS WHAT TO START WITH'
      $ 177 "Call Sub_AMR_MiR_V3"
      Sub_AMR_MiR_V3()
      $ 178 "get ugo data"
      $ 179 "Assign Tasks"
      $ 180 "TASK.ID = ugo_get_task()"
      TASK.ID = ugo_get_task()
      $ 181 "If TASK.ID≟1"
      if (TASK.ID == 1):
        $ 182 "Task_info≔'Charge'"
        global Task_info="Charge"
        $ 183 "Parameters"
        $ 184 "AMR_PosTarget≔1"
        global AMR_PosTarget=1
      else:
        $ 185 "ElseIf TASK.ID≟9"
        if (TASK.ID == 9):
          $ 186 "'Pick Sarstedt Rack from Variable source'"
          # 'Pick Sarstedt Rack from Variable source'
          $ 187 "Task_info≔'Navigate to Target'"
          global Task_info="Navigate to Target"
          $ 188 "Parameters"
          $ 189 "AMR_PosTarget≔UGO.read_input('00','ITM_ID')"
          global AMR_PosTarget=UGO.read_input("00","ITM_ID")
        else:
          $ 190 "ElseIf TASK.ID≟13"
          if (TASK.ID == 13):
            $ 191 "Task_info≔'Dose Powder'"
            global Task_info="Dose Powder"
            $ 192 "Parameters"
            $ 193 "ITM_ID≔1"
            global ITM_ID=1
            $ 194 "W_now≔(UGO.read_input('00','Container_weight'))/1000"
            global W_now=(UGO.read_input("00","Container_weight"))/1000
            $ 195 "Pow_name≔(UGO.read_input('00','Powder_name'))"
            global Pow_name=(UGO.read_input("00","Powder_name"))
            $ 196 "target_weight≔(UGO.read_input('00','Target_weight'))/1000"
            global target_weight=(UGO.read_input("00","Target_weight"))/1000
            $ 197 "send_picking_info(Pow_name,target_weight)"
            send_picking_info(Pow_name,target_weight)
            $ 198 "OBJ_Type≔6"
            global OBJ_Type=6
            $ 199 "JIG≔17"
            global JIG=17
            $ 200 "AMR_PosTarget≔5"
            global AMR_PosTarget=5
          else:
            $ 201 "ElseIf TASK.ID≟49"
            if (TASK.ID == 49):
              $ 202 "Task_info≔'Pick Containers'"
              global Task_info="Pick Containers"
              $ 203 "Parameters"
              $ 204 "ITM_ID≔1"
              global ITM_ID=1
              $ 205 "OBJ_Type≔6"
              global OBJ_Type=6
              $ 206 "JIG≔15"
              global JIG=15
              $ 207 "AMR_PosTarget≔3"
              global AMR_PosTarget=3
            else:
              $ 208 "ElseIf TASK.ID≟50"
              if (TASK.ID == 50):
                $ 209 "Task_info≔'Decap Containers'"
                global Task_info="Decap Containers"
                $ 210 "Parameters"
                $ 211 "ITM_ID≔1"
                global ITM_ID=1
                $ 212 "OBJ_Type≔6"
                global OBJ_Type=6
                $ 213 "JIG≔16"
                global JIG=16
                $ 214 "AMR_PosTarget≔5"
                global AMR_PosTarget=5
              else:
                $ 215 "ElseIf TASK.ID≟51"
                if (TASK.ID == 51):
                  $ 216 "Task_info≔'Detect Spatula and transfer powder'"
                  global Task_info="Detect Spatula and transfer powder"
                  $ 217 "Parameters"
                  $ 218 "ITM_ID≔1"
                  global ITM_ID=1
                  $ 219 "target_weight≔(UGO.read_input('00','Target_weight'))/1000"
                  global target_weight=(UGO.read_input("00","Target_weight"))/1000
                  $ 220 "OBJ_Type≔8"
                  global OBJ_Type=8
                  $ 221 "JIG≔16"
                  global JIG=16
                  $ 222 "AMR_PosTarget≔5"
                  global AMR_PosTarget=5
                else:
                  $ 223 "ElseIf TASK.ID≟52"
                  if (TASK.ID == 52):
                    $ 224 "Task_info≔'Pick Powder'"
                    global Task_info="Pick Powder"
                    $ 225 "Parameters"
                    $ 226 "ITM_ID≔1"
                    global ITM_ID=1
                    $ 228 "OBJ_Type≔6"
                    global OBJ_Type=6
                    $ 229 "JIG≔15"
                    global JIG=15
                    $ 230 "AMR_PosTarget≔3"
                    global AMR_PosTarget=3
                  else:
                    $ 231 "ElseIf TASK.ID≟53"
                    if (TASK.ID == 53):
                      $ 232 "Task_info≔'Decap Powder'"
                      global Task_info="Decap Powder"
                      $ 233 "Parameters"
                      $ 234 "ITM_ID≔1"
                      global ITM_ID=1
                      $ 235 "OBJ_Type≔6"
                      global OBJ_Type=6
                      $ 236 "JIG≔1"
                      global JIG=1
                      $ 237 "AMR_PosTarget≔5"
                      global AMR_PosTarget=5
                    else:
                      $ 238 "ElseIf TASK.ID≟54"
                      if (TASK.ID == 54):
                        $ 239 "Task_info≔'Empty and swap Powder container'"
                        global Task_info="Empty and swap Powder container"
                        $ 248 "Parameters"
                        $ 249 "ITM_ID≔1"
                        global ITM_ID=1
                        $ 251 "W_now≔(UGO.read_input('00','Container_weight'))/1000"
                        global W_now=(UGO.read_input("00","Container_weight"))/1000
                        $ 252 "Pow_name≔(UGO.read_input('00','Powder_name'))"
                        global Pow_name=(UGO.read_input("00","Powder_name"))
                        $ 255 "OBJ_Type≔6"
                        global OBJ_Type=6
                        $ 256 "JIG≔17"
                        global JIG=17
                        $ 257 "AMR_PosTarget≔5"
                        global AMR_PosTarget=5
                      else:
                        $ 258 "ElseIf TASK.ID≟55"
                        if (TASK.ID == 55):
                          $ 259 "Task_info≔'Place Powder'"
                          global Task_info="Place Powder"
                          $ 260 "Parameters"
                          $ 261 "ITM_ID≔1"
                          global ITM_ID=1
                          $ 262 "OBJ_Type≔6"
                          global OBJ_Type=6
                          $ 263 "JIG≔21"
                          global JIG=21
                          $ 264 "AMR_PosTarget≔5"
                          global AMR_PosTarget=5
                        else:
                          $ 265 "ElseIf TASK.ID≟56"
                          if (TASK.ID == 56):
                            $ 266 "Task_info≔'Dose Powder'"
                            global Task_info="Dose Powder"
                            $ 267 "Parameters"
                            $ 268 "ITM_ID≔1"
                            global ITM_ID=1
                            $ 269 "target_weight≔(UGO.read_input('00','Target_weight'))/1000"
                            global target_weight=(UGO.read_input("00","Target_weight"))/1000
                            $ 270 "W_now≔(UGO.read_input('00','Container_weight'))/1000"
                            global W_now=(UGO.read_input("00","Container_weight"))/1000
                            $ 271 "Pow_name≔(UGO.read_input('00','Powder_name'))"
                            global Pow_name=(UGO.read_input("00","Powder_name"))
                            $ 272 "OBJ_Type≔6"
                            global OBJ_Type=6
                            $ 273 "JIG≔17"
                            global JIG=17
                            $ 274 "AMR_PosTarget≔5"
                            global AMR_PosTarget=5
                          else:
                            $ 275 "ElseIf TASK.ID≟57"
                            if (TASK.ID == 57):
                              $ 276 "Task_info≔'Recipe Powder dosing'"
                              global Task_info="Recipe Powder dosing"
                              $ 277 "Parameters"
                              $ 278 "ITM_ID≔1"
                              global ITM_ID=1
                              $ 279 "Pow_A≔(UGO.read_input('00','PowderA'))"
                              global Pow_A=(UGO.read_input("00","PowderA"))
                              $ 280 "Pow_B≔(UGO.read_input('00','PowderB'))"
                              global Pow_B=(UGO.read_input("00","PowderB"))
                              $ 281 "Pow_C≔(UGO.read_input('00','PowderC'))"
                              global Pow_C=(UGO.read_input("00","PowderC"))
                              $ 282 "Total_weight≔(UGO.read_input('00','Total_weight'))/1000"
                              global Total_weight=(UGO.read_input("00","Total_weight"))/1000
                              $ 283 "Pow_A_percent≔(UGO.read_input('00','PowderA_percentage'))/100"
                              global Pow_A_percent=(UGO.read_input("00","PowderA_percentage"))/100
                              $ 284 "Pow_B_percent≔(UGO.read_input('00','PowderB_percentage'))/100"
                              global Pow_B_percent=(UGO.read_input("00","PowderB_percentage"))/100
                              $ 285 "Pow_C_percent≔(UGO.read_input('00','PowderC_percentage'))/100"
                              global Pow_C_percent=(UGO.read_input("00","PowderC_percentage"))/100
                              $ 286 "OBJ_Type≔6"
                              global OBJ_Type=6
                              $ 287 "JIG≔17"
                              global JIG=17
                              $ 288 "AMR_PosTarget≔5"
                              global AMR_PosTarget=5
                            else:
                              $ 289 "ElseIf TASK.ID≟58"
                              if (TASK.ID == 58):
                                $ 290 "Task_info≔'Pick Powder containers'"
                                global Task_info="Pick Powder containers"
                                $ 291 "Parameters"
                                $ 292 "ITM_ID≔1"
                                global ITM_ID=1
                                $ 293 "OBJ_Type≔6"
                                global OBJ_Type=6
                                $ 294 "JIG≔15"
                                global JIG=15
                                $ 295 "AMR_PosTarget≔3"
                                global AMR_PosTarget=3
                              else:
                                $ 296 "Else" "noBreak"
                                $ 297 "set_error(ERROR_WRONG_ORDER)"
                                set_error(ERROR_WRONG_ORDER)
                              end
                            end
                          end
                        end
                      end
                    end
                  end
                end
              end
            end
          end
        end
      end
      $ 298 "test ugo"
      $ 299 "Wait: 0.2"
      sleep(0.2)
      $ 300 "ugo_update_outputs()"
      ugo_update_outputs()
      $ 301 "If starting() and AMR_Done"
      if (starting()  and  AMR_Done):
        $ 302 "log_message(Task_info, 'New Task: ')"
        log_message(Task_info, "New Task: ")
        $ 303 "log_message(to_str(TASK.ID), 'Task_ID: ')"
        log_message(to_str(TASK.ID), "Task_ID: ")
        $ 304 "do_transition(keep_rxry=OBJ_Picked)"
        do_transition(keep_rxry=OBJ_Picked)
        $ 305 "STATE≔6"
        global STATE=6
        $ 306 "ugo_update_outputs()"
        ugo_update_outputs()
      end
    elif (6 == switch_1):
      $ 307 "Case 6"
      $ 308 "Execute"
      $ 309 "STATE_Info≔'Execute'"
      global STATE_Info="Execute"
      $ 310 "If  not CMD_Hold and not CMD_Suspend"
      global thread_flag_310=0
      thread Thread_if_310():
        $ 311 "Switch PROCESS_Step"
        switch_2 = PROCESS_Step
        $ 312 "Case 0"
        if (0 == switch_2):
          $ 313 "PROCESS_Info≔'process control'"
          global PROCESS_Info="process control"
          $ 314 "log_process(PROCESS_Info)"
          log_process(PROCESS_Info)
          $ 315 "process control"
          $ 316 "If  not AMR_AtTarget"
          if (  not  AMR_AtTarget):
            $ 317 "PROCESS_Step≔1"
            global PROCESS_Step=1
          else:
            $ 318 "ElseIf (( not ITM_Prepared and  not WRK_Done) or (ITM_Prepared and WRK_Done))"
            if (((  not  ITM_Prepared  and    not  WRK_Done)  or  (ITM_Prepared  and  WRK_Done))):
              $ 319 "PROCESS_Step≔2"
              global PROCESS_Step=2
            else:
              $ 320 "ElseIf  not WRK_Done"
              if (  not  WRK_Done):
                $ 321 "PROCESS_Step≔3"
                global PROCESS_Step=3
              else:
                $ 322 "Else" "noBreak"
                $ 323 "task finished"
                $ 324 "PROCESS_Info≔''"
                global PROCESS_Info=""
                $ 325 "STATE≔7"
                global STATE=7
                $ 326 "ugo_update_outputs()"
                ugo_update_outputs()
              end
            end
          end
        elif (1 == switch_2):
          $ 327 "Case 1"
          $ 328 "navigate"
          $ 329 "'MOVING THE uML'"
          # 'MOVING THE uML'
          $ 330 "PROCESS_Info≔'move to target'"
          global PROCESS_Info="move to target"
          $ 331 "log_process(PROCESS_Info)"
          log_process(PROCESS_Info)
          $ 332 "If TASK.ID≟1"
          if (TASK.ID == 1):
            $ 333 "Action≔51"
            global Action=51
          else:
            $ 334 "Else" "noBreak"
            $ 335 "Action≔52"
            global Action=52
          end
          $ 336 "Call Sub_AMR_MiR_V3"
          Sub_AMR_MiR_V3()
          $ 337 "If AMR_Done"
          if (AMR_Done):
            $ 338 "PROCESS_Step≔0"
            global PROCESS_Step=0
          end
        elif (2 == switch_2):
          $ 339 "Case 2"
          $ 340 "prepare"
          $ 341 "'THINGS THAT HAVE TO BE DONE ONCE IN A SEQUENCE,WORKFLOW'"
          # 'THINGS THAT HAVE TO BE DONE ONCE IN A SEQUENCE,WORKFLOW'
          $ 342 "PROCESS_Info≔'prepare for work'"
          global PROCESS_Info="prepare for work"
          $ 343 "log_process(PROCESS_Info)"
          log_process(PROCESS_Info)
          $ 344 "If TASK.WORK.ITM_ID_Src>1"
          if (TASK.WORK.ITM_ID_Src>1):
            $ 345 "ITM_ID≔TASK.WORK.ITM_ID_Src"
            global ITM_ID=TASK.WORK.ITM_ID_Src
          else:
            $ 346 "ElseIf TASK.WORK.ITM_ID_Tgt>1"
            if (TASK.WORK.ITM_ID_Tgt>1):
              $ 347 "ITM_ID≔TASK.WORK.ITM_ID_Tgt"
              global ITM_ID=TASK.WORK.ITM_ID_Tgt
            end
          end
          $ 348 "If  not ARM_Referenced and (ITM_ID≠0)"
          if (  not  ARM_Referenced  and  (ITM_ID != 0)):
            $ 349 "STP≔1"
            global STP=1
          else:
            $ 350 "ElseIf ARM_Referenced or (ITM_ID≟0)"
            if (ARM_Referenced  or  (ITM_ID == 0)):
              $ 351 "STP≔2"
              global STP=2
            end
          end
          $ 352 "Switch STP"
          switch_3 = STP
          $ 353 "Case 1"
          if (1 == switch_3):
            $ 354 "reference"
            $ 355 "STP_Info≔'reference at target position'"
            global STP_Info="reference at target position"
            $ 356 "log_step(STP_Info)"
            log_step(STP_Info)
            $ 357 "If ITM_ID≟1"
            if (ITM_ID == 1):
              $ 358 "CAM_Done≔ True "
              global CAM_Done=  True
            else:
              $ 359 "Else" "noBreak"
              $ 360 "Action≔131"
              global Action=131
              $ 361 "Call Sub_Vision_V18"
              Sub_Vision_V18()
            end
            $ 363 "If CAM_Done and  not ERROR.FLAG"
            if (CAM_Done  and    not  ERROR.FLAG):
              $ 364 "log_step('ARM referenced')"
              log_step("ARM referenced")
              $ 365 "ARM_Referenced≔ True "
              global ARM_Referenced=  True
            end
          elif (2 == switch_3):
            $ 366 "Case 2"
            $ 367 "manipulate"
            $ 368 "STP_Info≔'manipulate item'"
            global STP_Info="manipulate item"
            $ 369 "log_step(STP_Info)"
            log_step(STP_Info)
            $ 370 "'In case pressing button is needed'"
            # 'In case pressing button is needed'
            $ 371 "If found_in_list(ITM_ID, ITM_ID_List)"
            if (found_in_list(ITM_ID, ITM_ID_List)):
              $ 372 "Switch ITM_ID"
              switch_4 = ITM_ID
              $ 373 "Case 0"
              if (0 == switch_4):
                $ 374 "ITM_Manipulated≔ not ITM_Manipulated"
                global ITM_Manipulated=  not  ITM_Manipulated
              elif (1 == switch_4):
                $ 375 "Case 1"
                $ 376 "ITM_Manipulated≔ not ITM_Manipulated"
                global ITM_Manipulated=  not  ITM_Manipulated
              elif (2 == switch_4):
                $ 377 "Case 2"
              else:
                $ 387 "Default Case"
                $ 388 "ITM_Manipulated≔ not ITM_Manipulated"
                global ITM_Manipulated=  not  ITM_Manipulated
              end
            end
          end
          $ 389 "ITM_Prepared≔(ITM_Manipulated or  not found_in_list(ITM_ID, ITM_ID_List)) and (ARM_Referenced or ITM_ID≟0) and  not WRK_Done"
          global ITM_Prepared=(ITM_Manipulated  or    not  found_in_list(ITM_ID, ITM_ID_List))  and  (ARM_Referenced  or  ITM_ID == 0)  and    not  WRK_Done
          $ 390 "STP≔0"
          global STP=0
          $ 391 "STP_Info≔''"
          global STP_Info=""
          $ 392 "PROCESS_Step≔0"
          global PROCESS_Step=0
        elif (3 == switch_2):
          $ 393 "Case 3"
          $ 394 "work"
          $ 395 "'ADD EVERY MACHINE, OBJECT, STATION TO WORK ON'"
          # 'ADD EVERY MACHINE, OBJECT, STATION TO WORK ON'
          $ 396 "Switch ITM_ID"
          switch_3 = ITM_ID
          $ 397 "Case 1"
          if (1 == switch_3):
            $ 398 "uLM"
            $ 399 "If TASK.ID≟12"
            if (TASK.ID == 12):
              $ 400 "fill racks"
              $ 401 "Action≔151"
              global Action=151
              $ 402 "Call Sub_Vision_V18"
              Sub_Vision_V18()
              $ 403 "If  not ERROR.FLAG"
              if (  not  ERROR.FLAG):
                $ 404 "Actions for the task"
                $ 405 "Action≔1"
                global Action=1
                $ 406 "JIG≔2"
                global JIG=2
                $ 407 "JIG_Slot≔CAM_Result[0]"
                global JIG_Slot=CAM_Result[0]
                $ 408 "OBJ_Nbr≔CAM_Result[0]"
                global OBJ_Nbr=CAM_Result[0]
                $ 409 "OBJ_Type≔2"
                global OBJ_Type=2
                $ 410 "Call Sub_Action_V4"
                Sub_Action_V4()
                $ 411 "If OBJ_Picked"
                if (OBJ_Picked):
                  $ 412 "CAM_Result.remove(0)"
                  CAM_Result.remove(0)
                  $ 413 "PRC_TubCounter≔PRC_TubCounter+1"
                  global PRC_TubCounter=PRC_TubCounter+1
                  $ 414 "If PRC_TubCounter%4≟0"
                  if (PRC_TubCounter%4 == 0):
                    $ 415 "JIG_Slot≔4"
                    global JIG_Slot=4
                  else:
                    $ 416 "Else" "noBreak"
                    $ 417 "JIG_Slot≔PRC_TubCounter%4"
                    global JIG_Slot=PRC_TubCounter%4
                  end
                  $ 418 "OBJ_Nbr≔ceil(PRC_TubCounter/4)"
                  global OBJ_Nbr=ceil(PRC_TubCounter/4)
                  $ 419 "Action≔2"
                  global Action=2
                  $ 420 "JIG≔4"
                  global JIG=4
                  $ 421 "Call Sub_Action_V4"
                  Sub_Action_V4()
                  $ 422 "Action≔151"
                  global Action=151
                  $ 423 "Call Sub_Vision_V18"
                  Sub_Vision_V18()
                end
              end
              $ 424 "If (CAM_Captures≥CAM_PRM_Retries) or (PRC_TubCounter≥32)"
              if ((CAM_Captures >= CAM_PRM_Retries)  or  (PRC_TubCounter >= 32)):
                $ 425 "PROCESS_Step≔0"
                global PROCESS_Step=0
                $ 426 "WRK_Done≔ True "
                global WRK_Done=  True
              end
            else:
              $ 427 "ElseIf TASK.ID≟13"
              if (TASK.ID == 13):
                $ 428 "Dose Powder"
                $ 429 "Action≔131"
                global Action=131
                $ 430 "Call Sub_Vision_V18"
                Sub_Vision_V18()
                $ 431 "Action≔34"
                global Action=34
                $ 432 "Call Sub_Action_V4"
                Sub_Action_V4()
                $ 433 "PROCESS_Step≔0"
                global PROCESS_Step=0
                $ 434 "WRK_Done≔ True "
                global WRK_Done=  True
              else:
                $ 435 "ElseIf TASK.ID≟49"
                if (TASK.ID == 49):
                  $ 436 "Pick Powder container"
                  $ 437 "Action≔131"
                  global Action=131
                  $ 438 "Call Sub_Vision_V18"
                  Sub_Vision_V18()
                  $ 439 "Action≔35"
                  global Action=35
                  $ 440 "Call Sub_Action_V4"
                  Sub_Action_V4()
                  $ 441 "PROCESS_Step≔0"
                  global PROCESS_Step=0
                  $ 442 "WRK_Done≔ True "
                  global WRK_Done=  True
                else:
                  $ 443 "ElseIf TASK.ID≟50"
                  if (TASK.ID == 50):
                    $ 444 "Decap containers"
                    $ 445 "Action≔36"
                    global Action=36
                    $ 446 "Call Sub_Action_V4"
                    Sub_Action_V4()
                    $ 447 "PROCESS_Step≔0"
                    global PROCESS_Step=0
                    $ 448 "WRK_Done≔ True "
                    global WRK_Done=  True
                  else:
                    $ 449 "ElseIf TASK.ID≟51"
                    if (TASK.ID == 51):
                      $ 450 "Detect Spatula and transfer powder"
                      $ 451 "Action≔131"
                      global Action=131
                      $ 452 "Call Sub_Vision_V18"
                      Sub_Vision_V18()
                      $ 453 "Action≔37"
                      global Action=37
                      $ 454 "Call Sub_Action_V4"
                      Sub_Action_V4()
                      $ 455 "PROCESS_Step≔0"
                      global PROCESS_Step=0
                      $ 456 "WRK_Done≔ True "
                      global WRK_Done=  True
                    else:
                      $ 457 "ElseIf TASK.ID≟52"
                      if (TASK.ID == 52):
                        $ 458 "Pick Powder container"
                        $ 459 "Action≔131"
                        global Action=131
                        $ 460 "Call Sub_Vision_V18"
                        Sub_Vision_V18()
                        $ 461 "Action≔39"
                        global Action=39
                        $ 462 "Call Sub_Action_V4"
                        Sub_Action_V4()
                        $ 463 "PROCESS_Step≔0"
                        global PROCESS_Step=0
                        $ 464 "WRK_Done≔ True "
                        global WRK_Done=  True
                      else:
                        $ 465 "ElseIf TASK.ID≟53"
                        if (TASK.ID == 53):
                          $ 466 "Decap containerA"
                          $ 467 "Action≔40"
                          global Action=40
                          $ 468 "Call Sub_Action_V4"
                          Sub_Action_V4()
                          $ 469 "PROCESS_Step≔0"
                          global PROCESS_Step=0
                          $ 470 "WRK_Done≔ True "
                          global WRK_Done=  True
                        else:
                          $ 471 "ElseIf TASK.ID≟55"
                          if (TASK.ID == 55):
                            $ 472 "Place Powder"
                            $ 473 "Action≔131"
                            global Action=131
                            $ 474 "Call Sub_Vision_V18"
                            Sub_Vision_V18()
                            $ 475 "Action≔41"
                            global Action=41
                            $ 476 "Call Sub_Action_V4"
                            Sub_Action_V4()
                            $ 477 "PROCESS_Step≔0"
                            global PROCESS_Step=0
                            $ 478 "WRK_Done≔ True "
                            global WRK_Done=  True
                          else:
                            $ 479 "ElseIf TASK.ID≟54"
                            if (TASK.ID == 54):
                              $ 480 "Empty and swap container"
                              $ 481 "Action≔131"
                              global Action=131
                              $ 482 "Call Sub_Vision_V18"
                              Sub_Vision_V18()
                              $ 483 "Action≔42"
                              global Action=42
                              $ 484 "Call Sub_Action_V4"
                              Sub_Action_V4()
                              $ 485 "PROCESS_Step≔0"
                              global PROCESS_Step=0
                              $ 486 "WRK_Done≔ True "
                              global WRK_Done=  True
                            else:
                              $ 487 "ElseIf TASK.ID≟56"
                              if (TASK.ID == 56):
                                $ 488 "Dispense Powder"
                                $ 489 "Action≔131"
                                global Action=131
                                $ 490 "Call Sub_Vision_V18"
                                Sub_Vision_V18()
                                $ 491 "Action≔43"
                                global Action=43
                                $ 492 "Call Sub_Action_V4"
                                Sub_Action_V4()
                                $ 493 "PROCESS_Step≔0"
                                global PROCESS_Step=0
                                $ 494 "WRK_Done≔ True "
                                global WRK_Done=  True
                              else:
                                $ 495 "ElseIf TASK.ID≟57"
                                if (TASK.ID == 57):
                                  $ 496 "Recipe Dosing"
                                  $ 497 "Action≔48"
                                  global Action=48
                                  $ 498 "Call Sub_Action_V4"
                                  Sub_Action_V4()
                                  $ 515 "PROCESS_Step≔0"
                                  global PROCESS_Step=0
                                  $ 516 "WRK_Done≔ True "
                                  global WRK_Done=  True
                                else:
                                  $ 517 "ElseIf TASK.ID≟58"
                                  if (TASK.ID == 58):
                                    $ 518 "Pick Powder containers"
                                    $ 519 "Num_cont_picked≔0"
                                    global Num_cont_picked=0
                                    $ 520 "powder_position≔'Position1'"
                                    global powder_position="Position1"
                                    $ 521 "Loop Num_cont_picked<3"
                                    while (Num_cont_picked<3):
                                      $ 522 "Action≔131"
                                      global Action=131
                                      $ 523 "Call Sub_Vision_V18"
                                      Sub_Vision_V18()
                                      $ 524 "Action≔47"
                                      global Action=47
                                      $ 525 "Call Sub_Action_V4"
                                      Sub_Action_V4()
                                    end
                                    $ 526 "PROCESS_Step≔0"
                                    global PROCESS_Step=0
                                    $ 527 "WRK_Done≔ True "
                                    global WRK_Done=  True
                                  end
                                end
                              end
                            end
                          end
                        end
                      end
                    end
                  end
                end
              end
            end
          elif (2 == switch_3):
            $ 528 "Case 2"
          elif (5 == switch_3):
            $ 570 "Case 5"
          elif (20 == switch_3):
            $ 578 "Case 20"
          elif (43 == switch_3):
            $ 640 "Case 43"
          else:
            $ 648 "Default Case"
            $ 649 "WRK_Done≔ True "
            global WRK_Done=  True
            $ 650 "PROCESS_Step≔0"
            global PROCESS_Step=0
          end
        end
        thread_flag_310 = 1
      end
      if (  not  CMD_Hold and not CMD_Suspend):
        global thread_handler_310=run Thread_if_310()
        while (thread_flag_310 == 0):
          if not(  not  CMD_Hold and not CMD_Suspend):
            kill thread_handler_310
            thread_flag_310 = 2
          else:
            sync()
          end
        end
      else:
        thread_flag_310 = 2
      end
      $ 651 "If CMD_Hold"
      if (CMD_Hold):
        $ 652 "STATE≔9"
        global STATE=9
        $ 653 "ugo_update_outputs()"
        ugo_update_outputs()
      else:
        $ 654 "ElseIf CMD_Suspend"
        if (CMD_Suspend):
          $ 655 "STATE≔12"
          global STATE=12
          $ 656 "ugo_update_outputs()"
          ugo_update_outputs()
        end
      end
    elif (7 == switch_1):
      $ 657 "Case 7"
      $ 658 "Completing"
      $ 659 "STATE_Info≔'Completing'"
      global STATE_Info="Completing"
      $ 660 "'ADD COMMANDS FOR COMPLETING THE PROCESS'"
      # 'ADD COMMANDS FOR COMPLETING THE PROCESS'
      $ 661 "do_transition(keep_rxry=OBJ_Picked)"
      do_transition(keep_rxry=OBJ_Picked)
      $ 662 "Call Sub_AMR_MiR_V3"
      Sub_AMR_MiR_V3()
      $ 663 "If completing() and AMR_Done"
      if (completing()  and  AMR_Done):
        $ 664 "STATE≔8"
        global STATE=8
        $ 665 "ugo_update_outputs()"
        ugo_update_outputs()
      end
    elif (8 == switch_1):
      $ 666 "Case 8"
      $ 667 "Complete"
      $ 668 "STATE_Info≔'Complete'"
      global STATE_Info="Complete"
      $ 669 "If CMD_Reset"
      if (CMD_Reset):
        $ 670 "STATE≔3"
        global STATE=3
        $ 671 "ugo_update_outputs()"
        ugo_update_outputs()
      end
    elif (9 == switch_1):
      $ 672 "Case 9"
      $ 673 "Holding"
      $ 674 "STATE_Info≔'Holding'"
      global STATE_Info="Holding"
      $ 675 "stopl(0.5)"
      stopl(0.5)
      $ 676 "Call Sub_AMR_MiR_V3"
      Sub_AMR_MiR_V3()
      $ 677 "If holding() and AMR_Done"
      if (holding()  and  AMR_Done):
        $ 678 "STATE≔10"
        global STATE=10
        $ 679 "ugo_update_outputs()"
        ugo_update_outputs()
      end
    elif (10 == switch_1):
      $ 680 "Case 10"
      $ 681 "Held"
      $ 682 "STATE_Info≔'Held'"
      global STATE_Info="Held"
      $ 683 "If CMD_Unhold"
      if (CMD_Unhold):
        $ 684 "end_freedrive_mode()"
        end_freedrive_mode()
        $ 685 "STATE≔11"
        global STATE=11
        $ 686 "ugo_update_outputs()"
        ugo_update_outputs()
      else:
        $ 687 "ElseIf FNC_Freedrive"
        if (FNC_Freedrive):
          $ 688 "freedrive_mode()"
          freedrive_mode()
        else:
          $ 689 "Else" "noBreak"
          $ 690 "end_freedrive_mode()"
          end_freedrive_mode()
        end
      end
    elif (11 == switch_1):
      $ 691 "Case 11"
      $ 692 "Unholding"
      $ 693 "STATE_Info≔'Unholding'"
      global STATE_Info="Unholding"
      $ 694 "Clearing"
      $ 695 "Switch ERROR.ID"
      switch_2 = ERROR.ID
      $ 696 "Case 1002"
      if (1002 == switch_2):
        $ 697 "AMR_AtTarget≔ False "
        global AMR_AtTarget=  False
        $ 698 "ARM_Referenced≔ False "
        global ARM_Referenced=  False
        $ 699 "ITM_Prepared≔ False "
        global ITM_Prepared=  False
        $ 700 "PROCESS_Step≔1"
        global PROCESS_Step=1
      elif (2007 == switch_2):
        $ 701 "Case 2007"
        $ 702 "PROCESS_Step≔1"
        global PROCESS_Step=1
      end
      $ 703 "reset_error()"
      reset_error()
      $ 704 "reset_warning()"
      reset_warning()
      $ 705 "OBJ_Picked≔gripper_has_object()"
      global OBJ_Picked=gripper_has_object()
      $ 706 "Call Sub_AMR_MiR_V3"
      Sub_AMR_MiR_V3()
      $ 707 "If unholding() and AMR_Done"
      if (unholding()  and  AMR_Done):
        $ 708 "STATE≔6"
        global STATE=6
        $ 709 "ugo_update_outputs()"
        ugo_update_outputs()
      end
    elif (12 == switch_1):
      $ 710 "Case 12"
      $ 711 "Suspending"
      $ 712 "STATE_Info≔'Suspending'"
      global STATE_Info="Suspending"
      $ 713 "PROCESS_Info≔str_cat(PROCESS_Info, ' suspended')"
      global PROCESS_Info=str_cat(PROCESS_Info, " suspended")
      $ 714 "If suspending()"
      if (suspending()):
        $ 715 "STATE≔13"
        global STATE=13
        $ 716 "ugo_update_outputs()"
        ugo_update_outputs()
      end
    elif (13 == switch_1):
      $ 717 "Case 13"
      $ 718 "Suspended"
      $ 719 "STATE_Info≔'Suspended'"
      global STATE_Info="Suspended"
      $ 720 "Call Sub_AMR_MiR_V3"
      Sub_AMR_MiR_V3()
      $ 721 "If CMD_Unsuspend"
      if (CMD_Unsuspend):
        $ 722 "STATE≔14"
        global STATE=14
        $ 723 "ugo_update_outputs()"
        ugo_update_outputs()
      end
    elif (14 == switch_1):
      $ 724 "Case 14"
      $ 725 "Unsuspending"
      $ 726 "STATE_Info≔'Unsuspending'"
      global STATE_Info="Unsuspending"
      $ 727 "PROCESS_Step≔0"
      global PROCESS_Step=0
      $ 728 "If unsuspending()"
      if (unsuspending()):
        $ 729 "STATE≔6"
        global STATE=6
        $ 730 "ugo_update_outputs()"
        ugo_update_outputs()
      end
    elif (15 == switch_1):
      $ 731 "Case 15"
      $ 732 "Aborting"
      $ 733 "STATE_Info≔'Aborting'"
      global STATE_Info="Aborting"
      $ 734 "If aborting()"
      if (aborting()):
        $ 735 "STATE≔16"
        global STATE=16
        $ 736 "ugo_update_outputs()"
        ugo_update_outputs()
      end
    elif (16 == switch_1):
      $ 737 "Case 16"
      $ 738 "Aborted"
      $ 739 "STATE_Info≔'Aborted'"
      global STATE_Info="Aborted"
      $ 740 "If CMD_Clear"
      if (CMD_Clear):
        $ 741 "STATE≔17"
        global STATE=17
        $ 742 "ugo_update_outputs()"
        ugo_update_outputs()
      end
    elif (17 == switch_1):
      $ 743 "Case 17"
      $ 744 "Clearing"
      $ 745 "STATE_Info≔'Clearing'"
      global STATE_Info="Clearing"
      $ 746 "Clearing"
      $ 747 "reset_warning()"
      reset_warning()
      $ 748 "reset_error()"
      reset_error()
      $ 749 "If clearing()"
      if (clearing()):
        $ 750 "STATE≔2"
        global STATE=2
        $ 751 "ugo_update_outputs()"
        ugo_update_outputs()
      end
    end
    $ 752 "log_state(STATE_Info)"
    log_state(STATE_Info)
    $ 753 "log_warning(WARNING.MSG)"
    log_warning(WARNING.MSG)
    $ 754 "log_error(ERROR.MSG)"
    log_error(ERROR.MSG)
    $ 755 "Times"
    $ 756 "Switch STATE"
    switch_1 = STATE
    $ 757 "Case 1"
    if (1 == switch_1):
      $ 758 "TM_St_Stopping≔get_time(STATE_Times[STATE-1])"
      global TM_St_Stopping=get_time(STATE_Times[STATE-1])
    elif (2 == switch_1):
      $ 759 "Case 2"
      $ 760 "TM_St_Stopped≔get_time(STATE_Times[STATE-1])"
      global TM_St_Stopped=get_time(STATE_Times[STATE-1])
    elif (3 == switch_1):
      $ 761 "Case 3"
      $ 762 "TM_St_Resetting≔get_time(STATE_Times[STATE-1])"
      global TM_St_Resetting=get_time(STATE_Times[STATE-1])
    elif (4 == switch_1):
      $ 763 "Case 4"
      $ 764 "TM_St_Idle≔get_time(STATE_Times[STATE-1])"
      global TM_St_Idle=get_time(STATE_Times[STATE-1])
    elif (5 == switch_1):
      $ 765 "Case 5"
      $ 766 "TM_St_Starting≔get_time(STATE_Times[STATE-1])"
      global TM_St_Starting=get_time(STATE_Times[STATE-1])
    elif (6 == switch_1):
      $ 767 "Case 6"
      $ 768 "TM_St_Execute≔get_time(STATE_Times[STATE-1])"
      global TM_St_Execute=get_time(STATE_Times[STATE-1])
    elif (7 == switch_1):
      $ 769 "Case 7"
      $ 770 "TM_St_Completin≔get_time(STATE_Times[STATE-1])"
      global TM_St_Completin=get_time(STATE_Times[STATE-1])
    elif (8 == switch_1):
      $ 771 "Case 8"
      $ 772 "TM_St_Complete≔get_time(STATE_Times[STATE-1])"
      global TM_St_Complete=get_time(STATE_Times[STATE-1])
    elif (9 == switch_1):
      $ 773 "Case 9"
      $ 774 "TM_St_Holding≔get_time(STATE_Times[STATE-1])"
      global TM_St_Holding=get_time(STATE_Times[STATE-1])
    elif (10 == switch_1):
      $ 775 "Case 10"
      $ 776 "TM_St_Held≔get_time(STATE_Times[STATE-1])"
      global TM_St_Held=get_time(STATE_Times[STATE-1])
    elif (11 == switch_1):
      $ 777 "Case 11"
      $ 778 "TM_St_Unholding≔get_time(STATE_Times[STATE-1])"
      global TM_St_Unholding=get_time(STATE_Times[STATE-1])
    elif (12 == switch_1):
      $ 779 "Case 12"
      $ 780 "TM_St_Suspendin≔get_time(STATE_Times[STATE-1])"
      global TM_St_Suspendin=get_time(STATE_Times[STATE-1])
    elif (13 == switch_1):
      $ 781 "Case 13"
      $ 782 "TM_St_Suspended≔get_time(STATE_Times[STATE-1])"
      global TM_St_Suspended=get_time(STATE_Times[STATE-1])
    elif (14 == switch_1):
      $ 783 "Case 14"
      $ 784 "TM_St_Unsuspend≔get_time(STATE_Times[STATE-1])"
      global TM_St_Unsuspend=get_time(STATE_Times[STATE-1])
    elif (15 == switch_1):
      $ 785 "Case 15"
      $ 786 "TM_St_Aborting≔get_time(STATE_Times[STATE-1])"
      global TM_St_Aborting=get_time(STATE_Times[STATE-1])
    elif (16 == switch_1):
      $ 787 "Case 16"
      $ 788 "TM_St_Aborted≔get_time(STATE_Times[STATE-1])"
      global TM_St_Aborted=get_time(STATE_Times[STATE-1])
    elif (17 == switch_1):
      $ 789 "Case 17"
      $ 790 "TM_St_Clearing≔get_time(STATE_Times[STATE-1])"
      global TM_St_Clearing=get_time(STATE_Times[STATE-1])
    end
    $ 792 "Wait: 0.1"
    sleep(0.1)
  end
end
